(* IEC 61131-3 sources: llm-plc-st-eval/data/calibracion/gemini-3.1-pro-preview/B1/few_shot, 3 files *)

(* ---- ejec_1.st ---- *)
FUNCTION_BLOCK FB_Motor
VAR_INPUT
    btnMarcha : BOOL; (* Boton de marcha *)
    btnParo : BOOL; (* Boton de paro normal *)
    btnEmerg : BOOL; (* Boton de paro de emergencia *)
END_VAR
VAR_OUTPUT
    motorOn : BOOL; (* Activacion del motor *)
END_VAR
VAR
    trigMarcha : R_TRIG; (* Detector de flanco para evitar rearranque *)
END_VAR

(* Detecta nueva pulsacion de marcha para evitar rearranque si el boton sigue presionado *)
trigMarcha(CLK := btnMarcha);

(* Enclavamiento del motor con prioridad a las senales de paro *)
motorOn := (trigMarcha.Q OR motorOn) AND NOT btnParo AND NOT btnEmerg;
END_FUNCTION_BLOCK

(* ---- ejec_2.st ---- *)
FUNCTION_BLOCK FB_Motor
VAR_INPUT
    btnMarcha : BOOL; (* Boton de marcha *)
    btnParo : BOOL; (* Boton de paro *)
    btnEmerg : BOOL; (* Paro de emergencia *)
END_VAR
VAR_OUTPUT
    motorOn : BOOL; (* Estado del motor *)
END_VAR
VAR
    trigMarcha : R_TRIG; (* Detector de flanco de subida *)
END_VAR

(* Deteccion del flanco de subida para evitar rearranque si el boton sigue pulsado *)
trigMarcha(CLK := btnMarcha);

(* Control de arranque y paro con prioridad a las senales de detencion *)
motorOn := (trigMarcha.Q OR motorOn) AND NOT btnParo AND NOT btnEmerg;
END_FUNCTION_BLOCK

(* ---- ejec_3.st ---- *)
FUNCTION_BLOCK FB_Motor
VAR_INPUT
    btnMarcha : BOOL; (* Boton de marcha *)
    btnParo : BOOL;   (* Boton de paro *)
    btnEmerg : BOOL;  (* Paro de emergencia *)
END_VAR
VAR_OUTPUT
    motorOn : BOOL;   (* Estado del motor *)
END_VAR
VAR
    flancoMarcha : R_TRIG; (* Detector de flanco para evitar rearranque *)
END_VAR

(* Detectar flanco de subida para evitar rearranque si el boton sigue pulsado *)
flancoMarcha(CLK := btnMarcha);

(* Control de arranque y paro con prioridad a la detencion *)
IF btnParo OR btnEmerg THEN
    motorOn := FALSE;
ELSIF flancoMarcha.Q THEN
    motorOn := TRUE;
END_IF;
END_FUNCTION_BLOCK
